Fanuc KAREL source: kb00124.KL

-- PROVISIONAL review KL for V1013-1; original PC SHA256 0567c888947fa214841a1b3e3f756a69ef934c3ebda84373d6e0254741b6d131
-- Incomplete behavior may be omitted. Consult companion uncertainty JSON. Do not deploy.
PROGRAM KB00124
%NOLOCKGROUP
BEGIN
  -- UNRESOLVED_PC offsets 5-14; opcodes 3F,75
  -- UNRESOLVED_PC offsets 19-26; opcodes 9D,23
  -- UNRESOLVED_PC offsets 31-49; opcodes 27,22,2A,22,31
  -- UNRESOLVED_PC offsets 54-58; opcodes 7F
END KB00124
